// TIA Portal project "Clase3_PLCN3y4_ejercicio_variador_potenciometro_display" (V13)
// Uso de Norm, Escal y T_conv

(* hardware
DEVICE "S7-1200 station_1"  S7-1200 Station
   slot 0: "Rack_0"  Rack  V1.0
   slot 1: "PLC_1"  CPU 1214C AC/DC/Rly  6ES7 214-1BE30-0XB0  V2.2
   slot 3: "AQ 1x12BIT_1"  6ES7 232-4HA30-0XB0  V1.0
DEVICE "HMI_1"  KTP600 Basic color PN
   slot 0: "HMI"  HMI  6AV6 647-0AD11-3AX0  11.0.0.0
   slot 1: "HMI_RT_1"  KTP600 Basic color PN  6AV6 647-0AD11-3AX0  11.0.0.0
   slot 5: "HMI_1.IE_CP_1"  Interfaz PROFINET
      slot 1: "Interfaz PROFINET_1"  Interfaz PROFINET
         slot 1: "Port_1"  Port
*)

// ===== PLC "PLC_1"  CPU 1214C AC/DC/Rly =====

VAR_GLOBAL   // PLC tag table "Tabla de variables estándar"
   "hab" AT %I0.0 : Bool;
   "mem1" AT %M10.0 : Bool;
   "salida_hab" AT %Q0.0 : Bool;
   "value" AT %IW64 : UInt;
   "norm" AT %MD100 : Real;
   "scale" AT %MW120 : Word;
   "t_out" AT %MD220 : DWord;
   "sentido_giro" AT %Q0.1 : Bool;
   "Tag_1" AT %QW80 : Word;
   "abs_norm" AT %MW200 : Word;
END_VAR

ORGANIZATION_BLOCK "Main"   // OB1, LAD, ProgramCycle
TITLE = "Main Program Sweep (Cycle)"
{ S7_Optimized_Access := 'FALSE' }
VERSION : 0.1
BEGIN

REGION Network 1
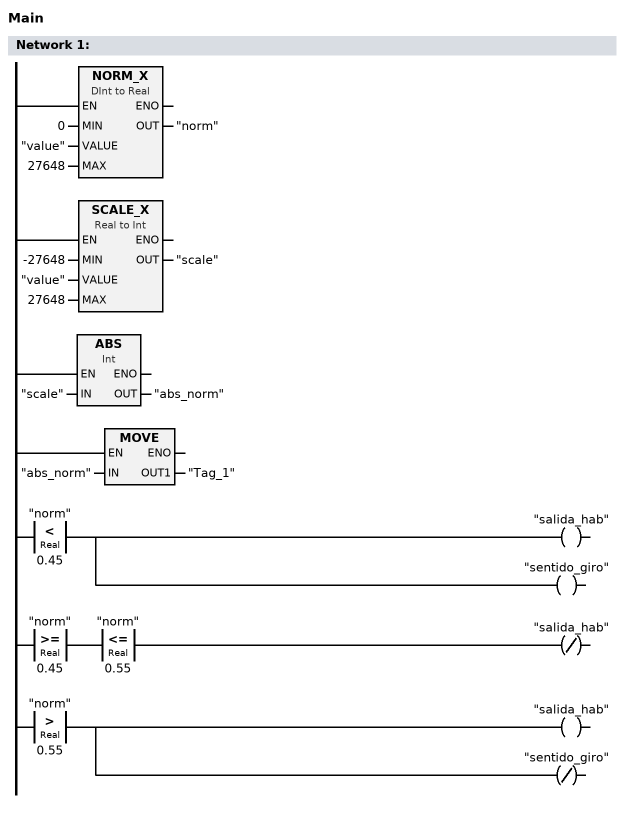
   RUNG wire#powerrail
      { S7_Templates := "[SrcType := DInt, DestType := Real]"; S7_GenerateENO := "TRUE" } Normalize(min := 0, value := "value", max := 27648, out => "norm")
   END_RUNG
   RUNG wire#powerrail
      { S7_Templates := "[SrcType := Real, DestType := Int]"; S7_GenerateENO := "TRUE" } Scale(min := -27648, value := "value", max := 27648, out => "scale")
   END_RUNG
   RUNG wire#powerrail
      { S7_Templates := "SrcType := Int"; S7_GenerateENO := "TRUE" } Abs(in := "scale", out => "abs_norm")
   END_RUNG
   RUNG wire#powerrail
      { S7_GenerateENO := "TRUE" } Move(in := "abs_norm", out1 => "Tag_1")
   END_RUNG
   RUNG wire#powerrail
      { S7_Templates := "SrcType := Real" } LT_Contact(in1 := "norm", in2 := 0.45)
      wire#w1
      Coil( "salida_hab" )
   END_RUNG
   RUNG wire#w1
      Coil( "sentido_giro" )
   END_RUNG
   RUNG wire#powerrail
      { S7_Templates := "SrcType := Real" } GE_Contact(in1 := "norm", in2 := 0.45)
      { S7_Templates := "SrcType := Real" } LE_Contact(in1 := "norm", in2 := 0.55)
      I_Coil( "salida_hab" )
   END_RUNG
   RUNG wire#powerrail
      { S7_Templates := "SrcType := Real" } GT_Contact(in1 := "norm", in2 := 0.55)
      wire#w2
      Coil( "salida_hab" )
   END_RUNG
   RUNG wire#w2
      I_Coil( "sentido_giro" )
   END_RUNG
   // the same network as SCL:
   "norm" := NORM_X(MIN := 0, VALUE := "value", MAX := 27648);
   "scale" := SCALE_X(MIN := -27648, VALUE := "value", MAX := 27648);
   "abs_norm" := ABS("scale");
   "Tag_1" := "abs_norm";
   "salida_hab" := "norm" < 0.45;
   "sentido_giro" := "salida_hab";
   "salida_hab" := NOT (("norm" >= 0.45) AND ("norm" <= 0.55));
   "salida_hab" := "norm" > 0.55;
   "sentido_giro" := NOT "salida_hab";
END_REGION
END_ORGANIZATION_BLOCK